(* IEC 61131-3 sources: PlcProgrammingProjects/Codesys4_Modbus/CodesysModbus.fbsdev/Application.iecapp^, 2 files *)

(* ---- modbus.gvl ---- *)
{attribute 'qualified_only'}
NAMESPACE modbus
VAR_GLOBAL

    now, currentIndex, counter, counter2 : INT;

    valueFromCodesys : INT;

    led1, led2, led3, led4 : BOOL;

    isAbove : BOOL;
END_VAR
END_NAMESPACE

(* ---- PLC_PRG.prg.st ---- *)
PROGRAM PLC_PRG
VAR
    counter : int ;
END_VAR

counter := counter + 1;

 modbus.valueFromCodesys :=  modbus.valueFromCodesys + 2;

 if modbus.valueFromCodesys > 100 then
      modbus.valueFromCodesys := 0;
 END_IF

END_PROGRAM
